(* IEC 61131-3 sources: IRIS-Project/LASAL CONTROL SOFTWARE/LasalProject_2025_09_25/Runtime/%LASALAPPDATA%/Runtime/Library/Loader/Source/code (part 11) *)

  retval := 1;

  IF (ops.tAbsolute - pUpdCell^.udLastUpdate) < (pUpdCell^.udUpdateRate AND 16#FFFF) THEN
    // udLastUpdate did not expire
    RETURN;
  END_IF;

  IF pUpdCell^.pCh = NIL THEN
    RETURN;
  END_IF;

  retval := 2;

  IF (pUpdCell^.udUpdateRate and UPDRATE_FLAG_IS_VBI) THEN
    dData := (pUpdCell^.pCh$^virtualBaseInit^.getCrc())$DINT;
  ELSIF (pUpdCell^.udUpdateRate AND UPDRATE_FLAG_IS_GLOBALVAR) THEN
//    dData := (pUpdCell^.pCh$^DINT)^;
    dData := UpDateGlobalVar(pUpdCell^.pCh, pUpdCell^.udUpdateRate);
  ELSE
    dData := rd(pUpdCell^.pCh);
  END_IF;

  IF dData = pUpdCell^.dData THEN
    // dData did not change
    pUpdCell^.udLastUpdate := ops.tAbsolute;
    RETURN;
  END_IF;

  retval := 3;

  // prepare the request message structure
  reqMsg.iOff  := iOff;
  reqMsg.pCh   := pUpdCell^.pCh;
  reqMsg.dData := dData;

  // Send the request
  rc := SendRequestR(pLogin,
                     CMD_UPDCELL,
                     respRequired:=FALSE,
                     pData:=#reqMsg,
                     dataLen:=SIZEOF(reqMsg),
                     blockingMode:=FALSE);
  IF rc <> 0 THEN
    DEBUG_VERBOSE2("%010d-*** UpdateCell(VarPos %d): SendCmdMsg failed, rc=%d", TO_UDINT(iOff), TO_UDINT(rc));
    // Dieser Fall tritt z.B. ein, wenn der Sendebuffer voll ist. Die Verbindung wird
    // nicht beendet, da die Zelle später auch noch übertragen werden kann, wenn wieder
    // Platz im Sendebuffer ist.
    retval := -rc;
  ELSE
    //DEBUGLOG2("%010d-UpdateCell: UPDCELL request sent, VarPos=%d, dData=0x%08X", TO_UDINT(iOff), TO_UDINT(dData));
    pUpdCell^.dData := dData;
    pUpdCell^.udLastUpdate := ops.tAbsolute;
  END_IF;

END_FUNCTION

//------------------------------------------------------------------------------
// UpdateListProcessorR
//------------------------------------------------------------------------------
FUNCTION UpdateListProcessorR
VAR_INPUT
  pLogin : ^loginContextR;
END_VAR
VAR
  list          : ^updateList;
  pUpdCell      : ^comStCell;  // pointer to cell in updatelist
  pStrtCell     : ^comStCell;
  rc : DINT;
END_VAR

  list := #pLogin^.statList;
  IF list^.nbrRefrCells > 0 THEN
    pStrtCell := list^.pActCell;
    WHILE 1 DO
      pUpdCell := list^.pActCell;

      rc := UpdateCellR(pLogin, pUpdCell, list^.actInd$UINT);
      IF rc <= 0 THEN
        RETURN;
      END_IF;

      IF (list^.actInd + 1) >= list^.nbrRefrCells THEN
        list^.actInd   := 0;
        list^.pActCell := list^.pFirstCell;
      ELSE
        list^.actInd   += 1;
        list^.pActCell += SIZEOF(list^.pActCell^);
      END_IF;

      IF pStrtCell = list^.pActCell THEN
        EXIT;
      END_IF;

      //Es wird nur 1 Zelle bei jedem Durchlauf gesendet, mehr macht bei
      //der seriellen Verbindung keinen Sinn.
      IF rc = 3 THEN
        EXIT;
      END_IF;
    END_WHILE;
  END_IF;

  list := #pLogin^.dynList;
  IF list^.nbrRefrCells > 0 THEN
    pStrtCell := list^.pActCell;
    WHILE 1 DO
      pUpdCell := list^.pActCell;

      rc := UpdateCellR(pLogin, pUpdCell, (list^.actInd + 1000)$UINT);
      IF rc <= 0 THEN
        RETURN;
      END_IF;

      IF (list^.actInd + 1) >= list^.nbrRefrCells THEN
        list^.actInd   := 0;
        list^.pActCell := list^.pFirstCell;
      ELSE
        list^.actInd   += 1;
        list^.pActCell += SIZEOF(list^.pActCell^);
      END_IF;

      IF pStrtCell = list^.pActCell THEN
        EXIT;
      END_IF;

      //Es wird nur 1 Zelle bei jedem Durchlauf gesendet, mehr macht bei
      //der seriellen Verbindung keinen Sinn.
      IF rc = 3 THEN
        EXIT;
      END_IF;
    END_WHILE;
  END_IF;

END_FUNCTION

//------------------------------------------------------------------------------
// SendAliveMessage_RS232
//------------------------------------------------------------------------------
FUNCTION SendAliveMessage_RS232
VAR_INPUT
  pLogin : ^loginContextR;
END_VAR
VAR_OUTPUT
    retval        : DINT;
END_VAR
VAR
    rc            : DINT;
END_VAR

  retval := 1;

  rc := SendRequestR(pLogin,
                     CMD_IAMALIVE,
                     respRequired:=FALSE,
                     pData:=NIL,
                     dataLen:=0,
                     blockingMode:=FALSE);
  IF rc <> 0 THEN
    DEBUGLOG1("%010d-*** SendAliveMessage_RS232: SendCmdMsg failed, rc=%d", TO_UDINT(rc));
    retval := rc;
  ELSE
    DEBUGLOG0("%010d-SendAliveMessage_RS232: IAMALIVE request sent");
  END_IF;

END_FUNCTION

//------------------------------------------------------------------------------
// SyncRefListsRS232
//  siehe Beschreibung von SyncRefLists
//------------------------------------------------------------------------------
FUNCTION SyncRefListsRS232
VAR_INPUT
  pLogin : ^loginContextR;
END_VAR
VAR
    obj     : pVoid;
    pHead   : ^IprHead;
    instr   : ^instruct;
END_VAR

#ifndef DUMMY_LOADER
    pHead := pLogin^.Com.GetHead();
#endif
    instr := pHead^.pCode;

    IF instr^.opCode = I_WRITE THEN

        obj := instr^.aPara[0]$^pVoid;

        // statische Refresh-Liste durchsuchen
        InvalidateRefListEntry(pLogin^.statList.pFirstCell, pLogin^.statList.nbrRefrCells$UINT, obj);

        // dynamische Refresh-Liste durchsuchen
        InvalidateRefListEntry(pLogin^.dynList.pFirstCell, pLogin^.dynList.nbrRefrCells$UINT, obj);

    END_IF;

END_FUNCTION

(*
  Stellt die MaxIdleTime ein
*)
FUNCTION SetMaxIdleTimeR
VAR_INPUT
  pLogin : ^loginContextR;
  maxIdleTime_ms : UDINT;
END_VAR

  IF maxIdleTime_ms <> pLogin^.maxIdleTime_ms THEN
    pLogin^.maxIdleTime_ms := maxIdleTime_ms;
    pLogin^.lastSendTime_ms := ops.tAbsolute - pLogin^.maxIdleTime_ms; // damit gleich was geschickt wird
  END_IF;

END_FUNCTION

(*
  ProcessCmdR
    Führt einen empfangenen Befehl aus.
*)
FUNCTION ProcessCmdR
VAR_INPUT
  pLogin : ^loginContextR;
  cmd : UINT;
  pData : pVoid;
  dataLen : UINT;
  pRespData : pVoid;
  pRespDataLen : ^UINT;
END_VAR
VAR_OUTPUT
  cmdProcessed : BOOL;
END_VAR
VAR
  bNext : UDINT;
  pResu : ^results;
  updList   : ^updateList;
  listType  : UDINT;
  pComCell  : ^comStCell;
  uiOffs    : UINT;
  data2LSE  : d2LSE;
  original_this : UDINT;
END_VAR

  cmdProcessed := FALSE;

  IF pLogin^.isClient THEN
    AliveCheckMsgRcvd(pLogin$^loginContext);
  END_IF;

  CASE cmd OF

    CMD_BEFIPR:
      DEBUGLOG1("%010d-~~~ ProcessCmd: BEFIPR, dataLen=%d", dataLen$UDINT);
      // req-data:
      //    workState   : iprStates;
      //    instr       : instruct;
      // resp-data:
      //    workState   : iprStates;
      //    resu        : results;
      cmdProcessed := TRUE;

      IF (dataLen < SIZEOF(iprStates)) | ((dataLen - SIZEOF(iprStates)) > SIZEOF(instruct)) THEN
        pRespData^$msgBefiprRespData.workstate := ERROR;
      ELSE
        // execute befipr
#ifndef DUMMY_LOADER
#ifdef LOADER_4_LASAL2
        _memcpy(pLogin^.com._m.head.pCode, #pData^$msgBefiprReqData.instr, dataLen - SIZEOF(iprStates));
        pLogin^.com._m.head.workstate := pData^$msgBefiprReqData.workstate;
        pLogin^.com._m.head.funkSt    := READY;
        pLogin^.com._m.resu.uilng :=0;
#else
        _memcpy(pLogin^.com.head.pCode, #pData^$msgBefiprReqData.instr, dataLen - SIZEOF(iprStates));
        pLogin^.com.head.workstate := pData^$msgBefiprReqData.workstate;
        pLogin^.com.head.funkSt    := READY;
        pLogin^.com.resu.uilng :=0;
#endif
        pRespData^$msgBefiprRespData.workstate := pLogin^.com.BEFIPR(#bNext);
#endif
        SyncRefListsRs232(pLogin);
      END_IF;

      // prepare the response
      pRespDataLen^ := SIZEOF(iprStates);
      IF pRespData^$msgBefiprRespData.workstate <> ERROR THEN
#ifndef DUMMY_LOADER
        pResu := pLogin^.com.GetResult();
#endif
        IF pResu^.uilng <> 16#FFFF THEN
          IF pResu^.uilng <= SIZEOF(pRespData^$msgBefiprRespData) THEN
            pRespDataLen^ += pResu^.uilng;
            _memcpy(#pRespData^$msgBefiprRespData.resu, pResu, pResu^.uilng);
          ELSE
#ifndef DUMMY_LOADER
#ifdef LOADER_4_LASAL2
            pLogin^.com._m.head.workstate := ERROR;
#else
            pLogin^.com.head.workstate := ERROR;
#endif
#endif
          END_IF;
        END_IF;
      END_IF;

    CMD_SESSINFO:
      DEBUGLOG1("%010d-~~~ ProcessCmd: SESSINFO, dataLen=%d", dataLen$UDINT);
      // req-data:
      //    version     : UDINT;
      // resp-data:
      //    version     : UDINT;

      IF dataLen >= (msgSessInfoData.sizeofDynList - msgSessInfoData.version) THEN

        cmdProcessed := TRUE;

        // prepare the response
        pRespDataLen^ := SIZEOF(msgSessInfoData);
        pRespData^$msgSessInfoData.version := COMLINKR_VERSION;
        pRespData^$msgSessInfoData.instId  := myInstanceID;
        pRespData^$msgSessInfoData.sessId  := 0;
        pRespData^$msgSessInfoData.sizeofDynList  := MAX_DYNLIST_ENTRIES;
        pRespData^$msgSessInfoData.sizeofStatList := MAX_STATLIST_ENTRIES;

#ifdef DEBUG
      ELSE
        DEBUG_VERBOSE0("%010d-~~~ ProcessCmd: dataLen too small");
#endif
      END_IF;

    CMD_TXUPD:
      DEBUGLOG2("%010d-~~~ ProcessCmd: CMD_TXUPD, dataLen=%d ofs=%d", dataLen$UDINT, TO_UDINT(pData^$msgTxUpdReqData.iOff));
      // req-data:
      //    iOff        : UINT;
      //    comcell     : comStCell;
      // resp-data:
      //    this request requires no response
      IF dataLen >= SIZEOF(msgTxUpdReqData) THEN

        cmdProcessed := TRUE;

        IF pData^$msgTxUpdReqData.iOff < 1000 THEN
          updList   := #pLogin^.statList;
          listType  := 0;
        ELSE
          updList   := #pLogin^.dynList;
          listType  := 1;
          pData^$msgTxUpdReqData.iOff -=1000;
        END_IF;

        IF TO_UDINT(pData^$msgTxUpdReqData.iOff) >= updList^.nbrCells THEN
          IF IncreaseUpdateList(updList, TO_UDINT(pData^$msgTxUpdReqData.iOff) + 1, listType) = NIL THEN
            DEBUGLOG0("%010d-*** ProcessCmd: MemoryUpdateList failed");
            DisconnectAfterErrorR(pLogin);
            RETURN;
          END_IF;
          DEBUGLOG2("%010d-*** ProcessCmd: updList %d increased to %d entries", listType, updList^.nbrCells);
        END_IF;

        pComCell := updList^.pFirstCell + (SIZEOF(comStCell) * pData^$msgTxUpdReqData.iOff);

        pComCell^ := pData^$msgTxUpdReqData.comcell;
        IF (pComCell^.udUpdateRate AND 0xFFFF) < SMALLEST_UPD_INTERVALL THEN
          pComCell^.udUpdateRate := (pComCell^.udUpdateRate AND 0xFFFF0000) OR SMALLEST_UPD_INTERVALL;
        END_IF;
        IF !!(pComCell^.udUpdateRate AND UPDRATE_FLAG_IS_GLOBALVAR) &
           GetdataBufferFlag(pComCell^.pCh$^VirtualBase) THEN
          // The object has the flag ATTR_DATA_BUFFER set. For these object more than
          // the 4 bytes of dData can be transmitted. The comlink server updates the cell
          // when the crc changes instead of dData.
          pComCell^.udUpdateRate := pComCell^.udUpdateRate or UPDRATE_FLAG_IS_VBI;
        END_IF;
#ifdef DEBUG
      ELSE
        DEBUG_VERBOSE0("%010d-~~~ ProcessCmd: dataLen too small");
#endif
      END_IF;

    CMD_SSREFR:
      DEBUGLOG2("%010d-~~~ ProcessCmd: SSREFR received, typ=%d, count=%d", TO_UDINT(pData^$msgSsRefrReqData.typ), TO_UDINT(pData^$msgSsRefrReqData.count));
      // req-data:
      //    count       : UINT;
      //    typ         : UINT;
      // resp-data:
      //    this request requires no response

      IF dataLen >= SIZEOF(msgSsRefrReqData) THEN

        cmdProcessed := TRUE;

        IF pData^$msgSsRefrReqData.typ = 0 THEN
          // static list
          LoadUpdateList(#pLogin^.statList, pData^$msgSsRefrReqData.count);
        ELSE
          // dynamic list
          LoadUpdateList(#pLogin^.dynList, pData^$msgSsRefrReqData.count);
        END_IF;
#ifdef DEBUG
      ELSE
        DEBUG_VERBOSE0("%010d-~~~ ProcessCmd: dataLen too small");
#endif
      END_IF;

    CMD_UPDCELL:
      DEBUGLOG2("%010d-~~~ ProcessCmd: UPDCELL received, dataLen=%d, VarPos=%d", dataLen$UDINT, TO_UDINT(pData^$msgUpdCellReqData.iOff));
      // req-data:
      //    iOff        : INT;
      //    comcell     : comStCell;
      // resp-data:
      //    this request requires no response

      IF dataLen >= SIZEOF(msgUpdCellReqData) THEN

        cmdProcessed := TRUE;

        uiOffs := pData^$msgUpdCellReqData.iOff$UINT;
        IF uiOffs < 1000 THEN
          pComCell := pLogin^.statList.pFirstCell;
          IF TO_UDINT(pData^$msgUpdCellReqData.iOff) >= pLogin^.statList.nbrCells THEN
            DEBUGLOG1("%010d-*** ProcessCmd: VarPos(%d) is too big for StatList", TO_UDINT(pData^$msgUpdCellReqData.iOff));
            RETURN;
          END_IF;
        ELSE
          uiOffs -=1000;
          pComCell := pLogin^.dynlist.pFirstCell;
          IF TO_UDINT(uiOffs) >= pLogin^.dynList.nbrCells THEN
            DEBUGLOG1("%010d-*** ProcessCmd: VarPos(%d) is too big for DynList", TO_UDINT(pData^$msgUpdCellReqData.iOff));
            RETURN;
          END_IF;
        END_IF;

        pComCell        := pComcell + (SIZEOF(comStCell) * uiOffs);

        IF pComCell^.pCh <> pData^$msgUpdCellReqData.pCh THEN
          DEBUGLOG0("%010d-*** ProcessCmd: invalid upd-cell received");
          RETURN;
        END_IF;
        pComCell^.dData := pData^$msgUpdCellReqData.dData;

        // call callback function
        IF pLogin^.pCallback <> NIL THEN
          data2LSE.data      := pComCell^.dData;
          data2LSE.uiOffs    := pData^$msgUpdCellReqData.iOff$UINT;
          data2LSE.varlistID := pComCell^.VarlistID;
          original_this := ESI;
          ESI := pLogin^.pThis;
          pLogin^.pCallback$PrototypeCallbackT(pLogin^.pComdefT, #data2LSE);
          ESI := original_this;
          DEBUG_VERBOSE3("%010d-~~~ ProcessCmd: Callback(dData=0x%08X,uiOffs=%d,id=0x%08X", TO_UDINT(data2LSE.data), TO_UDINT(data2LSE.uiOffs), TO_UDINT(data2LSE.varlistID));
        END_IF;
#ifdef DEBUG
      ELSE
        DEBUG_VERBOSE0("%010d-~~~ ProcessCmd: dataLen too small");
#endif
      END_IF;

    CMD_MAXIDLETIME:
      DEBUGLOG1("%010d-~~~ ProcessCmd: CMD_MAXIDLETIME received, maxIdleTime=%d", pData^$msgIdlTimReqData.maxIdleTime_ms);
      // req-data:
      //    maxIdleTime_ms : UDINT;
      // resp-data:
      //    this request requires no response

      cmdProcessed := TRUE;

      SetMaxIdleTimeR(pLogin, pData^$msgIdlTimReqData.maxIdleTime_ms);

    CMD_IAMALIVE:
      DEBUGLOG0("%010d-~~~ ProcessCmd: IAMALIVE received");
      // req-data:
      // resp-data:
      //    this request requires no response

      cmdProcessed := TRUE;

    CMD_LOGOUT:
      DEBUGLOG0("%010d-~~~ ProcessCmd: LOGOUT received");
      // req-data:
      //    this request requires no data
      // resp-data:
      //    this request requires no response
      LoadUpdateList( #pLogin^.statList, 0 );
      LoadUpdateList( #pLogin^.dynList, 0 );

    ELSE
      // unknown command
      DEBUGLOG2("%010d-~~~ ProcessCmd: unknown command received, cmd=0x%X, dataLen=%d", cmd$UDINT, dataLen$UDINT);

  END_CASE;

END_FUNCTION

(*
  ProcessCmdAndRespR
*)
FUNCTION ProcessCmdAndRespR
VAR_INPUT
  pLogin : ^loginContextR;
END_VAR
VAR
  pL1RecvBuffer : ^SER_L1_BUF;
  cmd : UINT;
  pData : pVoid;
  dataLen : UINT;
  respData : ARRAY[0..299] OF BYTE;
  respDataLen : UINT;
  seqNbr : UINT;
  ack : BOOL;
END_VAR

  pL1RecvBuffer := #pLogin^.rxL1BufReq;

  cmd := pL1RecvBuffer^.flagsCmd AND RS232_L1CMD_MASK;
  IF pL1RecvBuffer^.flagsCmd AND RS232_L1FLAGS_RESPONSE_REQUIRED THEN
    seqNbr := pL1RecvBuffer^.data$UINT;
    pData := #pL1RecvBuffer^.data[2];
    dataLen := pL1RecvBuffer^.dataLen - 2;
  ELSE
    pData := #pL1RecvBuffer^.data[0];
    dataLen := pL1RecvBuffer^.dataLen;
  END_IF;

  IF ProcessCmdR(pLogin, cmd, pData, dataLen, #respData[0], #respDataLen) THEN
    ack := TRUE;
  ELSE
    ack := FALSE;
  END_IF;

  IF pL1RecvBuffer^.flagsCmd AND RS232_L1FLAGS_RESPONSE_REQUIRED THEN
    SendResponseR(pLogin, seqNbr, ack, cmd, #respData[0], respDataLen);
  END_IF;

END_FUNCTION

(*
  Versucht, zu sendende Nodes aus der Queue zu entnehmen, in den L0-Buffer
  zu stellen, und den L0-Buffer dann zu schicken.
  Empfangene Daten werden in die Receive-Queue gestellt.

  Die Funktion blockiert nicht. Sie ist nicht thread-safe und wird daher nur
  aus dem Cyclic aufgerufen.
*)
FUNCTION ComlinkR_SerTransfer
VAR_INPUT
  pItf : ^RS232_ITF;
END_VAR
VAR_OUTPUT
  event : BOOL;
END_VAR
VAR
  pL0RecvBuffer : ^SER_L0_BUF;
  nextOfs : UDINT;
  nRead : UDINT;
  pL1Buffer : ^SER_L1_BUF;
  dstChIdx : UDINT;
  pLogin : ^loginContextR; // connection context
  flags : BYTE;
END_VAR

  event := FALSE;

  LOCK_R();
  IF pItf^.bytesToSend = 0 THEN
    // Es gibt dzt. nichts zu senden, daher im L0SendBufferCollect nachschauen,
    // ob Daten vorhanden sind oder ob der Timeout für die anstehende Response
    // abgelaufen ist.
    IF (pItf^.pL0SendBufferCollect^.dataLen > L0_EMPTY_DATALEN) |
       (pItf^.l0RespNecessary & (ops.tAbsolute - pItf^.l0RespNecessaryTimeval_ms)$DINT > 0)
    THEN
      // Es soll was gesendet werden.
      // -> L0SendBufferCollect auf den anderen Buffer umschalten und das
      // Senden anstossen, indem bytesToSend auf >0 gesetzt wird.
      pItf^.pL0SendBufferCollect := SwitchL0Buffer(pItf, pItf^.pL0SendBufferCollect);
      pItf^.bytesToSend := pItf^.pL0SendBufferTransfer^.dataLen + L0_EMPTY_DATALEN;
      pItf^.bytesSent := 0;
      DEBUGLOG1("%010d-    SerTransfer: L0 send data available, bytesToSend: %d", TO_UDINT(pItf^.bytesToSend));
      OS_MT_Pulse(comlinkEventR);
      event := TRUE;
    END_IF;
  END_IF;

  IF pItf^.bytesToSend > 0 THEN
    // Es gibt was zu senden.
    IF !!pItf^.sendInProgress THEN
      L0CheckSend(pItf);
    END_IF;
    IF pItf^.sendInProgress THEN
      L0Send(pItf);
    END_IF;
    IF pItf^.bytesToSend = 0 THEN
      // Es konnte alles gesendet werden
      // -> Den L0SendBufferTransfer so vorbereiten, dass er wieder Daten aufsammeln
      // kann und dann L0SendBufferTransfer auf den anderen Buffer umschalten.
      IF pItf^.pL0SendBufferTransfer^.flagsCmd AND RS232_L0FLAGS_IS_REQUEST THEN
        // es ist ein Request gesendet worden, daher ist ab jetzt eine Response anstehend
        pItf^.l0RespPending := TRUE;
        pItf^.l0RespPendingTimeout_ms := ops.tAbsolute + pItf^.timeoutVal;
      ELSE
        // es ist eine Response gesendet worden, daher ist ab jetzt keine mehr anstehend,
        pItf^.l0RespNecessary := FALSE;
      END_IF;
      pItf^.pL0SendBufferTransfer^.dataLen := L0_EMPTY_DATALEN;
      pItf^.pL0SendBufferTransfer := SwitchL0Buffer(pItf, pItf^.pL0SendBufferTransfer);
      pItf^.sendInProgress := FALSE;
      DEBUGLOG2("%010d->>> SerTransfer: L0 finished send, new flags: respPending=%d, respNecessary=%d", pItf^.l0RespPending, pItf^.l0RespNecessary);
    END_IF;
  END_IF;

  pL0RecvBuffer := L0Recv(pItf);
  UNLOCK_R();

  IF pL0RecvBuffer <> NIL THEN
    DEBUGLOG1("%010d-<<< SerTransfer: L0 received data, datlen=%d", pL0RecvBuffer^.dataLen);
    nextOfs := SER_L0_BUF.data;
    WHILE nextOfs < (pL0RecvBuffer^.dataLen + 2) DO
      pL1Buffer := ScanL1Block(pL0RecvBuffer, #nextOfs, #nRead);
      flags := pL1Buffer^.flagsCmd AND (RS232_L1FLAGS_IS_REQUEST OR
                                        RS232_L1FLAGS_RESPONSE_REQUIRED);
      IF flags = (RS232_L1FLAGS_IS_REQUEST OR RS232_L1FLAGS_RESPONSE_REQUIRED) THEN
        // Es handelt sich um einen Request, der beantwortet werden möchte.
        DEBUGLOG2("%010d-<1  SerTransfer: got L1 Request that needs a response, dst=%d, src=%d", TO_UDINT(pL1Buffer^.dstChIdx), TO_UDINT(pL1Buffer^.srcChIdx));
        dstChIdx := pL1Buffer^.dstChIdx;
        IF (dstChIdx < 255) & (loginArrayR[dstChIdx] <> NIL) THEN
          DEBUG_VERBOSE0("%010d-*** SerTransfer: processing command");
          pLogin := loginArrayR[dstChIdx];
          _memcpy(#pLogin^.rxL1BufReq, pL1Buffer, nRead);
          ProcessCmdAndRespR(pLogin);
        ELSIF dstChIdx = 255 &
              GetL1CmdR(pL1Buffer) = CMD_CONNECT &
              pL1Buffer^.dataLen >= 2 THEN
          DEBUGLOG0("%010d-*** SerTransfer: processing login");
          // es will sich jemand einloggen
          pLogin := SearchUsedConnBlockSvrR(pItf^.itfIdx, pL1Buffer^.srcChIdx);
          IF pLogin = NIL THEN
            pLogin := AllocNewConnBlockSvrR(pItf^.itfIdx, pL1Buffer^.srcChIdx);
            DEBUGLOG2("%010d-    SerTransfer: allocated new channel, myChIdx=%d, hisChIdx=%d", pLogin^.myChIdx, pLogin^.hisChIdx);
          ELSE
            DEBUGLOG2("%010d-    SerTransfer: re-using old channel, myChIdx=%d, hisChIdx=%d", pLogin^.myChIdx, pLogin^.hisChIdx);
          END_IF;
          IF pLogin <> NIL THEN
            ResetL1(pLogin);
            // Die MaxIdleTime wird auf einen Wert <> 0 gesetzt, damit der Server
            // die Verbindung abbricht, wenn keine Kommunikation mehr stattfindet.
            // Das ist bei RS232 wichtig, weil sich ja um eine temporäre Modemverbindung
            // handeln könnte.
            SetMaxIdleTimeR(pLogin, 10000(*10Sek.*));

            pLogin^.hisChIdx := pL1Buffer^.srcChIdx;
            pLogin^.isConnected := TRUE;
#ifndef DUMMY_LOADER
            pLogin^.Com.InitCode(FALSE);
#endif
            SendResponseR(pLogin,
                          GetL1SeqNbrR(pL1Buffer),
                          ack := TRUE,
                          pL1Buffer^.flagsCmd AND RS232_L1CMD_MASK,
                          pData := NIL,
                          dataLen := 0);
          END_IF;

        END_IF;
      ELSIF flags = RS232_L1FLAGS_IS_REQUEST THEN
        DEBUGLOG2("%010d-<1  SerTransfer: got L1 Request, dst=%d, src=%d", TO_UDINT(pL1Buffer^.dstChIdx), TO_UDINT(pL1Buffer^.srcChIdx));
        dstChIdx := pL1Buffer^.dstChIdx;
        IF (dstChIdx < 255) & (loginArrayR[dstChIdx] <> NIL) THEN
          DEBUG_VERBOSE0("%010d-*** SerTransfer: processing command");
          pLogin := loginArrayR[dstChIdx];
          _memcpy(#pLogin^.rxL1BufReq, pL1Buffer, nRead);
          ProcessCmdAndRespR(pLogin);
        END_IF;
      ELSE
        // Es handelt sich um eine Response
        DEBUGLOG2("%010d-    SerTransfer: got L1 Response, dst=%d, src=%d", TO_UDINT(pL1Buffer^.dstChIdx), TO_UDINT(pL1Buffer^.srcChIdx));
        dstChIdx := pL1Buffer^.dstChIdx;
        IF (dstChIdx < 255) & (loginArrayR[dstChIdx] <> NIL) THEN
          pLogin := loginArrayR[dstChIdx];
          IF GetL1CmdR(pL1Buffer) = CMD_CONNECT THEN
            pLogin^.hisChIdx := pL1Buffer^.srcChIdx;
          END_IF;
          IF pL1Buffer^.srcChIdx = pLogin^.hisChIdx THEN
            DEBUGLOG0("%010d-    SerTransfer: finish pending response");
            _memcpy(#pLogin^.rxL1BufResp.dstChIdx, pL1Buffer + 1, nRead - 1);
            // Wenn srcChIdx im L1 RxBuffer auf <>INVALID_CHIDX gesetzt wird, dann heisst das,
            // dass der Buffer voll ist und vom Aufrufer ausgewertet werden darf.
            pLogin^.rxL1BufResp.srcChIdx := pL1Buffer^$BYTE;
            OS_MT_Pulse(comlinkEventR);
            event := TRUE;
          ELSE
            DEBUGLOG0("%010d-*** SerTransfer: no pending response in this channel");
            DisconnectAfterErrorR(pLogin);
          END_IF;
        END_IF;
      END_IF;
    END_WHILE;
  END_IF;

END_FUNCTION

//------------------------------------------------------------------------------
// ComlinkR_CyWork
//------------------------------------------------------------------------------
FUNCTION ComlinkR_CyWork
VAR
  i : UDINT;
  pLogin : ^loginContextR; // connection context
  pItf : ^RS232_ITF;
END_VAR

  IF !!g_RS232activity THEN
    // Aus Performancegründen wird hier gleich zurückgesprungen, wenn keiner
    // eine RS232 Kommunikation anfgefordert hat.
    RETURN;
  END_IF;

  FOR i := 0 TO arraysize(rs232Itfs)-1 DO
    pItf := #rs232Itfs[i];
    IF pItf^.hComm <> 0 THEN
      IF pItf^.fnInitInterface <> NIL THEN
        // Callback Funktion aufrufen, damit die Anwendung die Möglichkeit hat, eine
        // Modemverbindung zu beenden
        IF pItf^.fnInitInterface$LDR_InitRs232Interface(
              pItf^.pThis, ComlinkR_Idx2Itfnbr(i$DINT), pItf^.hCommAppl) <= 0 THEN
          LOCK_R();
          pItf^.hComm := 0;
          UNLOCK_R();
          EXIT;
        END_IF;
      END_IF;
      ComlinkR_SerTransfer(pItf);

      // Wenn das RespPending Flag länger als l0RespPendingTimeout_ms ansteht,
      // dann ist wahrscheinlich die Gegenstation nicht mehr aktiv.
      IF pItf^.l0RespPending & ((ops.tAbsolute - pItf^.l0RespPendingTimeout_ms)$DINT > 0) THEN
        DEBUGLOG0("%010d-*** ComlinkR_CyWork: timeout for l0RespPending exceeded, resetting itf");
        DisconnectAllForItf(pItf);
        ResetL0(pItf);
      END_IF;

    ELSIF pItf^.startServer THEN
      pItf^.hComm := ComlinkR_GetHandle(ComlinkR_Idx2Itfnbr(i$DINT));
    END_IF;
  END_FOR;

  FOR i := 0 TO (arraysize(loginArrayR) - 1) DO
    pLogin := loginArrayR[i];
    IF pLogin <> NIL & !!pLogin^.isClient THEN
      IF IsConnectedR(pLogin) THEN
        IF pLogin^.txL1BufCmd.dataValid THEN
          // Es gibt eine Response, die wegen zu wenig Platz im L0 Buffer
          // noch nicht gesendet werden konnte
          LOCK_R();
          PackL1Block(pLogin, #pLogin^.txL1BufCmd);
          UNLOCK_R();
        END_IF;

        UpdateListProcessorR(pLogin);

        IF pLogin^.maxIdleTime_ms > 0 THEN
          IF ops.tAbsolute - pLogin^.lastSendTime_ms > pLogin^.maxIdleTime_ms THEN
            SendAliveMessage_RS232(pLogin); // der Gegenstelle mitteilen, daß man noch lebt
          END_IF;
        END_IF;
      END_IF;
    END_IF;
  END_FOR;

END_FUNCTION

(*
  Diese Funktion wird von der Anwendung aufgerufen, wenn entweder die
  Standardeinstellungen der RS232 Schnittstelle verändert werden sollen,
  oder wenn der Loader einen Server auf einer RS232 Schnittstelle aktivieren
  soll.
  Der Server ist auf einer RS232 Schnittstelle standardmäßig nicht aktiv,
  weil sonst wären alle verfügbaren RS232 Schnittstellen vom Loader belegt.
*)
FUNCTION GLOBAL __CDECL LDR_SetRs232ComlinkParams
VAR_INPUT
  interface : UDINT;
  baudrate : UINT;
  startServer : DINT;
  fnInitInterface : pVoid;
  pThis : pVoid;
END_VAR
VAR_OUTPUT
  retVal : DINT;
END_VAR
VAR
  idx : DINT;
END_VAR

  retVal := 0;

  idx := ComlinkR_Itfnbr2Idx(interface);

  IF idx >= 0 THEN
    IF baudrate <> 16#FFFF THEN
      rs232Itfs[idx].baudrate := baudrate;
      rs232Itfs[idx].timeoutVal := GetL0TimeoutValR(rs232Itfs[idx].baudrate);
      DEBUGLOG2("%010d-    LDR_SetRs232ComlinkParams: itf %d - timeoutVal=%d", idx$UDINT, rs232Itfs[idx].timeoutVal);
    END_IF;
    IF startServer <> -1 THEN
      rs232Itfs[idx].startServer := startServer;
      g_RS232activity := TRUE;
    END_IF;
    IF fnInitInterface <> NIL THEN
      rs232Itfs[idx].fnInitInterface := fnInitInterface;
      rs232Itfs[idx].pThis := pThis;
    END_IF;
  ELSE
    retVal := -1;
  END_IF;

END_FUNCTION

VAR_GLOBAL
  aSoc          : ARRAY [0..63] OF DINT;
END_VAR

#ifdef LOADER_TCP_MODERATE
FUNCTION TCPIP_Task
VAR_INPUT
  pvoid       : ^void;
END_VAR
VAR
  i           : DINT;
  SocNum      : DINT;
  aSocPtr     : ARRAY [0..63] OF ^bufferedsocket;
  pLogin      : ^loginContext;
  pCmdConn    : ^cmdConnBlock;
  pRefrConn   : ^refrConnBlock;
END_VAR

  while 1 do
    OS_MT_DELAY(5);

    //--------------------------------------------------------------------
    // reset the number of sockets
    //--------------------------------------------------------------------
    SocNum := 0;

    //--------------------------------------------------------------------
    // T C P   C L I E N T   S O C K E T S
    //--------------------------------------------------------------------
    if (loginanz) then
      for i := 0 to (g_max_logins - 1) do
        pLogin := loginarray[i];
        if (pLogin <> NIL) then
          aSoc[SocNum] := pLogin^.refrSockClnt.sock;
          aSocPtr[SocNum] := #pLogin^.refrSockClnt;
          SocNum += 1;
        end_if;
      end_for;
    end_if;

    //--------------------------------------------------------------------
    // T C P   C O M M A N D   S E R V E R   S O C K E T S
    //--------------------------------------------------------------------
    if (nbrCmdConn) then
      pCmdConn := pCmdConnRoot;
      while (pCmdConn <> NIL) do
        aSoc[SocNum] := pCmdConn^.bsock.sock;
        aSocPtr[SocNum] := #pCmdConn^.bsock;
        SocNum += 1;
        pCmdConn := pCmdConn^.next;
      end_while;
    end_if;

    //--------------------------------------------------------------------
    // T C P   R E F R E S H   S E R V E R   S O C K E T S
    //--------------------------------------------------------------------
    if (nbrRefrConn) then
      pRefrConn := pRefrConnRoot;
      while (pRefrConn <> NIL) do
        aSoc[SocNum] := pRefrConn^.bsock.sock;
        aSocPtr[SocNum] := #pRefrConn^.bsock;
        SocNum += 1;
        pRefrConn := pRefrConn^.next;
      end_while;
    end_if;

    //--------------------------------------------------------------------
    // // look for available data
    //--------------------------------------------------------------------
    if (SocNum) then
      OS_TCP_USER_SELECT(SocNum,                  // Anzahl der Sockets
                         #aSoc[0],                // Pointer auf Socket-Array
                         SELECT_OPT_READ,         // Option
                         0,                       // Flag -> wird
                         0);

      for i := 0 to (SocNum - 1) do
        if (aSoc[i] > 0) then
          aSocPtr[i]$^bufferedsocket^.isDataAvailable := true;
        end_if;
      end_for;
    end_if;

  end_while;

END_FUNCTION
#endif

#endif // COMLINK_LASAL
